(*
SPDX-FileCopyrightText: © 2026 Oleksandr Tiutyk <trofimich@gmail.com>
SPDX-License-Identifier: MIT
License: https://opensource.org/license/mit
*)

(*!
<summary>Runs one multi-cycle test until completion or the inherited deadline.</summary>
<description>
Map this program to one cyclic PLC task or call its Execute method once per cycle from that task.
The concrete runner owns the tests; the program owns the reporter and performs task
cleanup at the end of every scan. Inspect _Runner.IsFinished, AllPassed and counts, then _Report.IsReady.
For independent task execution, assign SingleCycleTestExample and MultiCycleTestExample to different tasks.
They share no instances or mutable buffers. Do not assign the same program instance to multiple tasks.
</description>
*)

{attribute 'no_explicit_call' := 'do not call this function block directly'}
PROGRAM MultiCycleTestExample
VAR
	{attribute 'hide'}
	_ClassName : STRING := __POUNAME();

	_Runner : TimerDelayTestRunner;
	_Report : TOF_Testing.JUnitXmlReporter;
	_Configured : BOOL;
END_VAR

Execute();

//! <summary>Borrows the concrete program name for its lifetime; callers must not modify it.</summary>
{attribute 'monitoring' := 'call'}
PROPERTY ClassName : REFERENCE TO STRING
GET
ClassName REF= _ClassName;
END_GET
END_PROPERTY

(*!
<summary>Advances this example and performs standalone task-boundary memory cleanup.</summary>
<description>
Call once per cycle from the owning task, either through this method or by mapping this PROGRAM to that task.
Do not drive both entry paths or share the instance between tasks. Use as the standalone example in its task;
hosts with additional transient-exception consumers must provide a shared boundary instead.
</description>
*)
METHOD Execute
IF NOT _Configured THEN
	_Runner.Reporter := _Report;
	_Configured := TRUE;
END_IF

_Runner.Execute(cleanupTaskMemory := TRUE);
END_METHOD

(*!
<summary>Provides the library namespace used in diagnostics.</summary>
<description>
Borrowed read-only reference to the compiler-initialized library namespace; no ownership transfer.
</description>
*)
{attribute 'monitoring' := 'call'}
PROPERTY NamespaceName : REFERENCE TO STRING
GET
NamespaceName REF= CurrentNamespace.Name;
END_GET
END_PROPERTY

END_PROGRAM

(* stored: Version 1.1.0.1
   POU MultiCycleTestExample: Id {833032c1-474b-4136-851b-0270f1d7109d}, SpecialFunc None
   Property ClassName: Id {3634cb61-f6a6-4a16-b98a-c4a8acf3fd64}
   Get Get: Id {b9b0cbd4-b141-434d-85b6-8634754ea93a}
   Method Execute: Id {772e4cb0-483f-43da-984f-ceb595d0d3aa}
   Property NamespaceName: Id {2b6075ee-6ecb-4842-8b33-7b3bc9a3b693}
   Get Get: Id {7ea4fd38-93c9-466c-ab52-31a9c96c663e} *)
